(* IEC 61131-3 sources: Testing02/Test_Version_Control/Temp/Import/TS_Test_UT/Logical/TS_UnitTest/Libraries/UtMgr, 3 files *)

(* ---- UtMgr.typ ---- *)
(********************************************************************
 * COPYRIGHT -- Bernecker + Rainer
 ********************************************************************
 * Library: UtMgr
 * File: UtMgr.typ
 * Author: B+R
 ********************************************************************
 * Data types of library UtMgr
 ********************************************************************)

TYPE
	UtMgrLocationType : 	STRUCT  (*Provides location information as passed by a assert*)
		TestSetName : UDINT; (*&STRING Name of current Test Set*)
		TestCaseName : UDINT; (*&STRING Name of current Test Case*)
		Line : UDINT; (*Line number (utMgrTEST_TYPE_C)*)
		Location : UDINT; (*&STRING Location information *)
		File : UDINT; (*&STRING File name*)
	END_STRUCT;
	UtMgrInformationalType : 	STRUCT  (*Informational Data, will be reset before test run is active*)
		TestCasesSinceActiveCounter : UDINT; (*Counts executed test cases (increments at the beginning of a test case)*)
		FailedAssertCounter : UDINT; (*Counts total failed asserts since start of testsuite execution *)
		PassedAssertCounter : UDINT; (*Counts total passed asserts since start of testsuite execution *)
		InformationalMessageCounter : UDINT; (*Counts total informational messages since start of testsuite execution *)
		LastKnownPassedLocation : UtMgrLocationType; (*Provides information about last known location (as reported in a test assert)*)
	END_STRUCT;
	UtMgrTestTypeEnum :
		( (*Defines Implementation of  UtMgrTestSuite*)
		utMgrTEST_TYPE_NONE := 0, (*Invalid value*)
		utMgrTEST_TYPE_C := 10, (*Test Suite uses the static library UnitTest *)
		utMgrTEST_TYPE_OTHER := 20 (*Reserved*)
		);
	UtMgrTestPhaseBasicHelperEnum :
		( (*Internal status of test execution*)
		utMgrTEST_PHASE_IDLE := 0, (*No tests running*)
		utMgrTEST_PHASE_RUNNING := 5, (*Executing Test Sets*)
		utMgrTEST_PHASE_DONE := 10 (*Done executing Test Sets*)
		);
	UtMgrUnitTestRunnerHelperType : 	STRUCT  (*Internal*)
		TestSets : UDINT; (*Pointer to the array of Test Sets*)
		TestSetCount : UINT; (*Number of entries in array*)
		CurrentPhase : UtMgrTestPhaseBasicHelperEnum; (*Status of internal test execution*)
		CurrentTestSet : UINT; (*Index of current active Test Set*)
	END_STRUCT;
	UtMgrSuiteInternalType : 	STRUCT  (*Internal*)
		State : DINT; (*Internal*)
		Handle : UDINT; (*Internal*)
		List : ARRAY[0..29]OF UDINT; (*Internal*)
		LibInst : UDINT; (*Internal*)
		TestHelper : UtMgrUnitTestRunnerHelperType; (*Internal*)
	END_STRUCT;
END_TYPE

(* ---- UtMgr.fun ---- *)
(********************************************************************
 * COPYRIGHT -- Bernecker + Rainer
 ********************************************************************
 * Library: UtMgr
 * File: UtMgr.fun
 * Author: B+R
 ********************************************************************
 * Functions and function blocks of library UtMgr
 ********************************************************************)

FUNCTION_BLOCK UtMgrTestSuite (*Represents a test suite*)
	VAR_INPUT
		Enable : BOOL; (*Enables FB*)
		Name : STRING[80]; (*Distinct name of test suite*)
		Description : STRING[200]; (*Description of the test suite*)
		Type : UtMgrTestTypeEnum; (*Type of test suite*)
		MetaInformation : STRING[200]; (*Meta information. Data will be copied to the report at the end of the test suite execution*)
		TestAborted : BOOL; (*Rising edge = Test aborted*)
		TestFinished : BOOL; (*Rising edge = Test finished*)
	END_VAR
	VAR_OUTPUT
		Busy : BOOL; (*FB is busy*)
		Active : BOOL; (*FB is active*)
		Error : BOOL; (*Indicates an error*)
		StatusID : DINT; (*Status information*)
		TestActive : BOOL; (*Test suite  is active*)
		Informational : UtMgrInformationalType; (*Monitoring information*)
		TestFinishedAck : BOOL; (*Acknowledge of flag "TestFinished"*)
		TestFinishedDone : BOOL; (*Test suite finished, report is done*)
	END_VAR
	VAR
		Internal : UtMgrSuiteInternalType;
	END_VAR
END_FUNCTION_BLOCK

FUNCTION_BLOCK UtMgrMonitor (*Provides diagnostic data for monitoring*)
	VAR_INPUT
		Enable : BOOL; (*Enables FB*)
	END_VAR
	VAR_OUTPUT
		Active : BOOL; (*FB is active*)
		Error : BOOL; (*Indicates an error*)
		StatusID : DINT; (*Status information*)
		TestActive : BOOL; (*A test suite is active*)
		Informational : UtMgrInformationalType; (*Informational data provided while FB is active*)
	END_VAR
END_FUNCTION_BLOCK

FUNCTION UtMgrTestRunnerRunTest : DINT (*Internal: Used by the static library UnitTest. Handles Test Set execution*)
	VAR_INPUT
		TestSet : UDINT; (*&TestSet*)
	END_VAR
END_FUNCTION

(* ---- UtMgr.var ---- *)
(********************************************************************
 * COPYRIGHT -- Bernecker + Rainer
 ********************************************************************
 * Library: UtMgr
 * File: UtMgr.var
 * Author: B+R
 ********************************************************************
 * Constants of library UtMgr
 ********************************************************************)
VAR CONSTANT
	utERR_GENERAL : DINT := -1057750784; (*General error, see help*)
	utMgrERR_INVALID_PARAM : DINT := -1057750783; (*Check parameters*)
	utMgrERR_TOO_MANY_TESTS : DINT := -1057750782; (*Too many UtMgrTestSuites enabled, disable unused instances*)
END_VAR
